FUNCTION_BLOCK LampControl (* CAT Function Block Type *)
  (* Standard: 61499-2 *)
  (* Version 0.0, 8/3/2026, template *)
  PACKAGE Main;
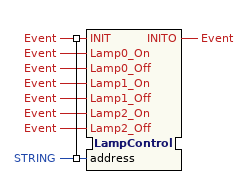
  EVENT_INPUT
    INIT WITH address; (* Initialization Request *)
    Lamp0_On; (* Normal Execution Request *)
    Lamp0_Off;
    Lamp1_On;
    Lamp1_Off;
    Lamp2_On;
    Lamp2_Off;
  END_EVENT
  EVENT_OUTPUT
    INITO; (* Initialization Confirm *)
  END_EVENT
  VAR_INPUT
    address : STRING; (* Input event qualifier *)
  END_VAR
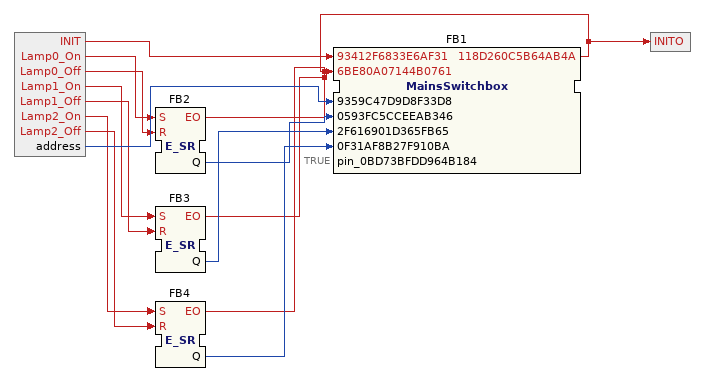
  FBS
    FB1 : MainsSwitchbox(pin_0BD73BFDD964B184 := TRUE);
    FB2 : E_SR;
    FB3 : E_SR;
    FB4 : E_SR;
  END_FBS
  EVENT_CONNECTIONS
    FB1.118D260C5B64AB4A TO INITO;
    Lamp2_On TO FB4.S;
    Lamp2_Off TO FB4.R;
    Lamp1_On TO FB3.S;
    Lamp1_Off TO FB3.R;
    Lamp0_On TO FB2.S;
    Lamp0_Off TO FB2.R;
    INIT TO FB1.93412F6833E6AF31;
    FB1.118D260C5B64AB4A TO FB1.6BE80A07144B0761;
    FB2.EO TO FB1.6BE80A07144B0761;
    FB3.EO TO FB1.6BE80A07144B0761;
    FB4.EO TO FB1.6BE80A07144B0761;
  END_CONNECTIONS
  DATA_CONNECTIONS
    address TO FB1.9359C47D9D8F33D8;
    FB2.Q TO FB1.0593FC5CCEEAB346;
    FB3.Q TO FB1.2F616901D365FB65;
    FB4.Q TO FB1.0F31AF8B27F910BA;
  END_CONNECTIONS
END_FUNCTION_BLOCK
